(* Logix 5000 project; controller R400_500_XLS vendor 1 type 14 code 216 rev 31.11; software revision 31.01; part 20 of 32 *)
(* tags used below, declared in another part *)
   Alarm : SINT;   // Wait 3 seconds
   AlarmAcked : BOOL;   // Alarm has been acked
   AlarmFlag : DINT;   // Active alarm flag
   AlarmFlag1 : DINT;
   AlarmMuted : BOOL;
   AlarmTran0 : BOOL;   // Transition from step 3 to step 0
   Ashutdown : SINT;   // Not Used
   bAlrm : BOOL[64];
   Critical_Alarm : BOOL;
   CycExcBuffer : UDT_CYCLE;
   F2rinse : DINT;   // Not Used
   F3rinse : DINT;   // Not Used
   FC45_NextMaintDate : DINT[3];   // Next maintenance due date
   FINALRINSE_1 : DINT;   // Final rinse 1 id number
   HeatSmp : DINT;
   I_0_Missing : BOOL;
   L310ER_Led : DINT;
   LowPressAlmSp : REAL;   // Pump pressure too low setpoint
   M : DINT[5];   // Memory Bits
   ONS_FC45 : DINT;
   PWTnkTempAlmSp : REAL;   // Pure water tank temperature too high setpoint
   ResetMute : BOOL;
   Run : DINT;
   SumpTempAlmSp : REAL;   // Sump temperature too high setpoint
   Supervisor : DINT;
   Tmr : TIMER[107];
   Trt_Wsh : DINT;
   AlarmAck : INT;   // Alarm acknowledgement from the HMI
   AlarmTrigger : INT;   // Triggers the alarm screen if different of 0
   BatteryLowWarning : BOOL;
   bONSAuditTrailAlarm : BOOL;
   Current_Screen : DINT;
   DateTime : DINT[7];
   FC45_NbCycBeforeMaint : DINT;
   I_Ld_Dr_Cls_Sw : BOOL;   // Load door close
   I_MCR : BOOL;   // MCR input
   I_Mtr_Ovrld : BOOL;   // Motor overload
   I_Pw_Tnk_Sft_Lvl_Sw : BOOL;   // Pure water tank safety level switch
   I_Smp_Sft_Lvl_Sw : BOOL;   // Sump safety level switch
   I_Unld_Dr_Cls_Sw : BOOL;   // Unload door close
   I_UnldDr_ClseSlnce_Bttn : BOOL;   // Door Close/ Silence button Unload Side
   LastRecircSumpDrainTemp : REAL;
   Load : Doors;
   LoadDoorClosing : BOOL;
   LoadDoorOpening : BOOL;
   PmpPres : REAL;
   PureWaterTankTemp : REAL;   // Pure water tank temperature
   PWT_DeltaTempNeg : REAL;
   PWT_DeltaTempPos : REAL;
   Screen_Ctrl : DINT;   // PLC Screen Request
   SimGenEnabled : BOOL;   // SimGen enable bit 1= Simgen ON
   SPV_19 : BOOL;   // Screen 80 Enabled/Disabled Pump pressure monitoring
   SumpTemp : REAL;   // Sump temperature in °C
   tDelayBeforeFillingAuthAlarm : TIMER;
   tDelayBeforeTankFillingAuthAlarm : TIMER;
   Tpb : DINT[11];
   TreatmentPtr : DINT;
   udtAuditTrail : UDT_AuditTrail;
   Unit : Hrdwre;   // Unit Configuration
   UnLoad : Doors;
   UnloadDoorClosing : BOOL;
   UnloadDoorOpening : BOOL;
(* MainProgram, continued *)

ROUTINE WSH_10_WSH_37_GENERATE_ALARM_DISPLAY   (* ladder *)
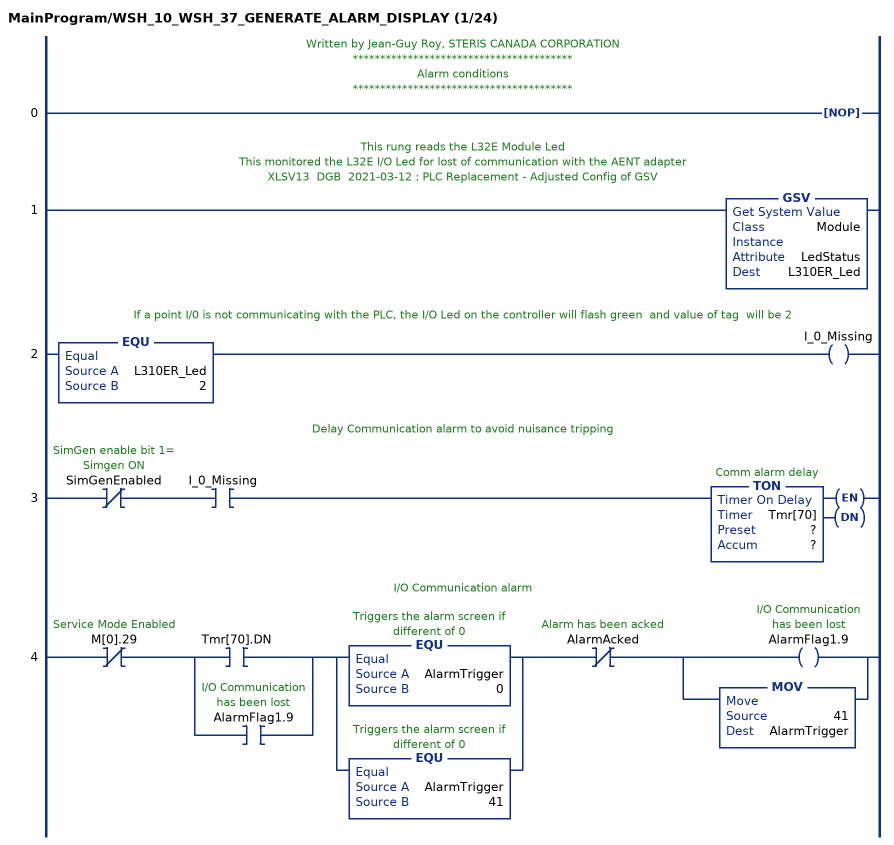
   // Written by Jean-Guy Roy, STERIS CANADA CORPORATION
   // ****************************************
   // Alarm conditions
   // ****************************************
   0: NOP();
   // This rung reads the L32E Module Led
   // This monitored the L32E I/O Led for lost of communication with the AENT adapter
   // XLSV13  DGB  2021-03-12 : PLC Replacement - Adjusted Config of GSV
   1: GSV(Module,,LedStatus,L310ER_Led);
   // If a point I/0 is not communicating with the PLC, the I/O Led on the controller will flash green  and value of tag  will be 2
   2: EQU(L310ER_Led,2)OTE(I_0_Missing);
   // Delay Communication alarm to avoid nuisance tripping
   3: XIO(SimGenEnabled)XIC(I_0_Missing)TON(Tmr[70],?,?);
   // I/O Communication alarm
   4: XIO(M[0].29)[XIC(Tmr[70].DN) ,XIC(AlarmFlag1.9) ][EQU(AlarmTrigger,0) ,EQU(AlarmTrigger,41) ]XIO(AlarmAcked)[OTE(AlarmFlag1.9) ,MOV(41,AlarmTrigger) ];
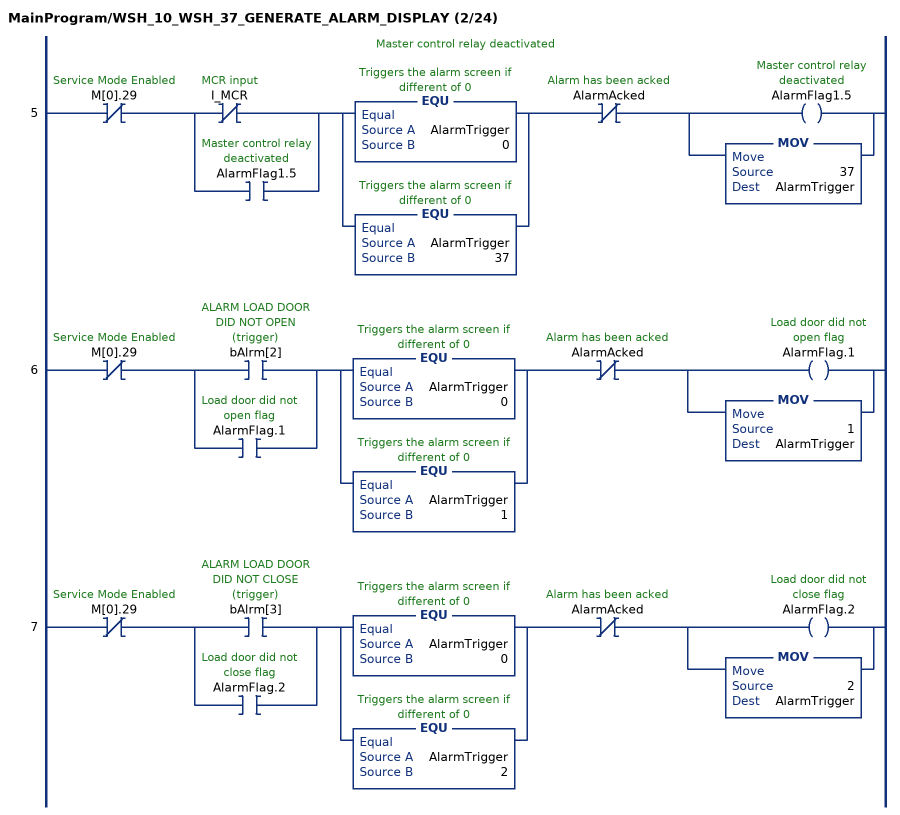
   // Master control relay deactivated
   5: XIO(M[0].29)[XIO(I_MCR) ,XIC(AlarmFlag1.5) ][EQU(AlarmTrigger,0) ,EQU(AlarmTrigger,37) ]XIO(AlarmAcked)[OTE(AlarmFlag1.5) ,MOV(37,AlarmTrigger) ];
   6: XIO(M[0].29)[XIC(bAlrm[2]) ,XIC(AlarmFlag.1) ][EQU(AlarmTrigger,0) ,EQU(AlarmTrigger,1) ]XIO(AlarmAcked)[OTE(AlarmFlag.1) ,MOV(1,AlarmTrigger) ];
   7: XIO(M[0].29)[XIC(bAlrm[3]) ,XIC(AlarmFlag.2) ][EQU(AlarmTrigger,0) ,EQU(AlarmTrigger,2) ]XIO(AlarmAcked)[OTE(AlarmFlag.2) ,MOV(2,AlarmTrigger) ];
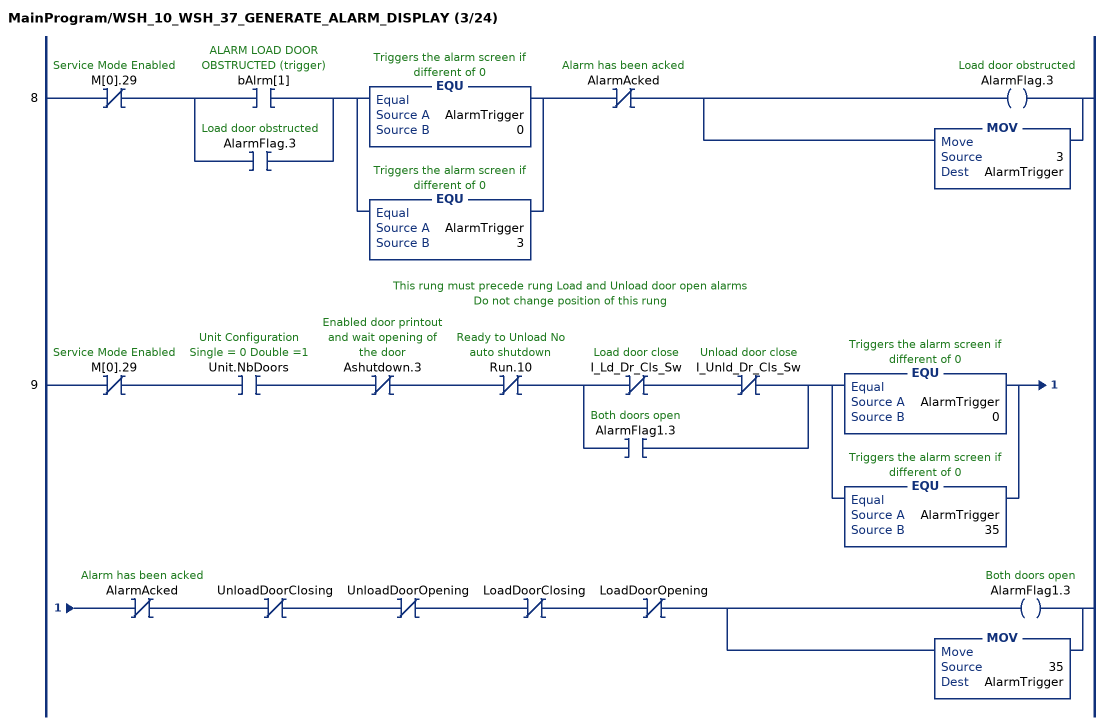
   8: XIO(M[0].29)[XIC(bAlrm[1]) ,XIC(AlarmFlag.3) ][EQU(AlarmTrigger,0) ,EQU(AlarmTrigger,3) ]XIO(AlarmAcked)[OTE(AlarmFlag.3) ,MOV(3,AlarmTrigger) ];
   // This rung must precede rung Load and Unload door open alarms
   // Do not change position of this rung
   9: XIO(M[0].29)XIC(Unit.NbDoors)XIO(Ashutdown.3)XIO(Run.10)[XIO(I_Ld_Dr_Cls_Sw) XIO(I_Unld_Dr_Cls_Sw) ,XIC(AlarmFlag1.3) ][EQU(AlarmTrigger,0) ,EQU(AlarmTrigger,35) ]XIO(AlarmAcked)XIO(UnloadDoorClosing)XIO(UnloadDoorOpening)XIO(LoadDoorClosing)XIO(LoadDoorOpening)[OTE(AlarmFlag1.3) ,MOV(35,AlarmTrigger) ];
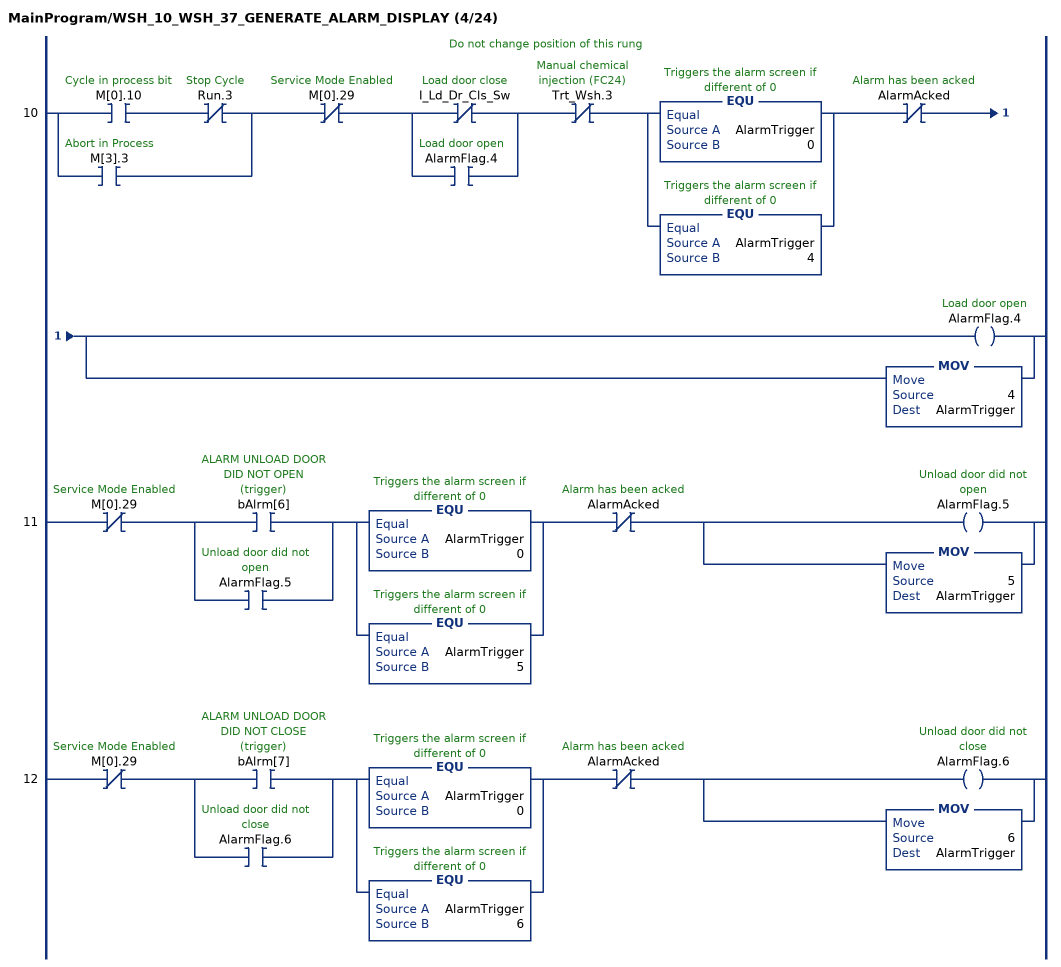
   // Do not change position of this rung
   10: [XIC(M[0].10) XIO(Run.3) ,XIC(M[3].3) ]XIO(M[0].29)[XIO(I_Ld_Dr_Cls_Sw) ,XIC(AlarmFlag.4) ]XIO(Trt_Wsh.3)[EQU(AlarmTrigger,0) ,EQU(AlarmTrigger,4) ]XIO(AlarmAcked)[OTE(AlarmFlag.4) ,MOV(4,AlarmTrigger) ];
   11: XIO(M[0].29)[XIC(bAlrm[6]) ,XIC(AlarmFlag.5) ][EQU(AlarmTrigger,0) ,EQU(AlarmTrigger,5) ]XIO(AlarmAcked)[OTE(AlarmFlag.5) ,MOV(5,AlarmTrigger) ];
   12: XIO(M[0].29)[XIC(bAlrm[7]) ,XIC(AlarmFlag.6) ][EQU(AlarmTrigger,0) ,EQU(AlarmTrigger,6) ]XIO(AlarmAcked)[OTE(AlarmFlag.6) ,MOV(6,AlarmTrigger) ];
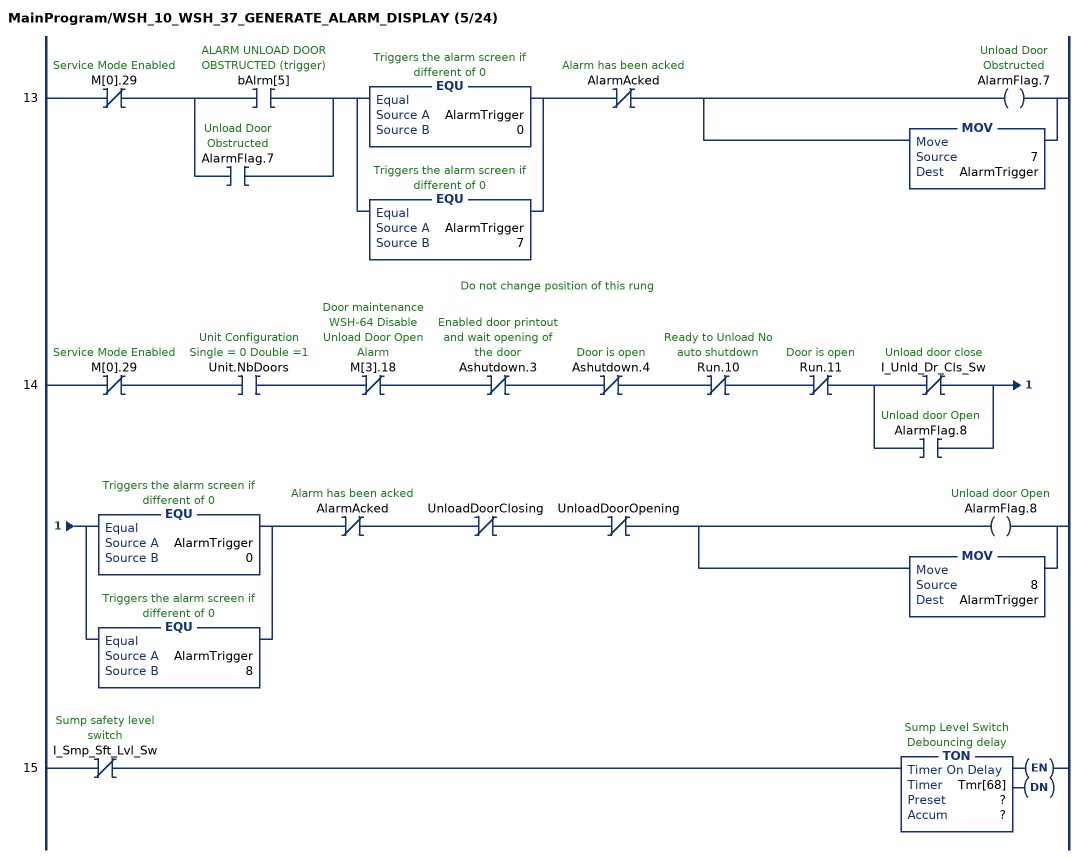
   13: XIO(M[0].29)[XIC(bAlrm[5]) ,XIC(AlarmFlag.7) ][EQU(AlarmTrigger,0) ,EQU(AlarmTrigger,7) ]XIO(AlarmAcked)[OTE(AlarmFlag.7) ,MOV(7,AlarmTrigger) ];
   // Do not change position of this rung
   14: XIO(M[0].29)XIC(Unit.NbDoors)XIO(M[3].18)XIO(Ashutdown.3)XIO(Ashutdown.4)XIO(Run.10)XIO(Run.11)[XIO(I_Unld_Dr_Cls_Sw) ,XIC(AlarmFlag.8) ][EQU(AlarmTrigger,0) ,EQU(AlarmTrigger,8) ]XIO(AlarmAcked)XIO(UnloadDoorClosing)XIO(UnloadDoorOpening)[OTE(AlarmFlag.8) ,MOV(8,AlarmTrigger) ];
   15: XIO(I_Smp_Sft_Lvl_Sw)TON(Tmr[68],?,?);
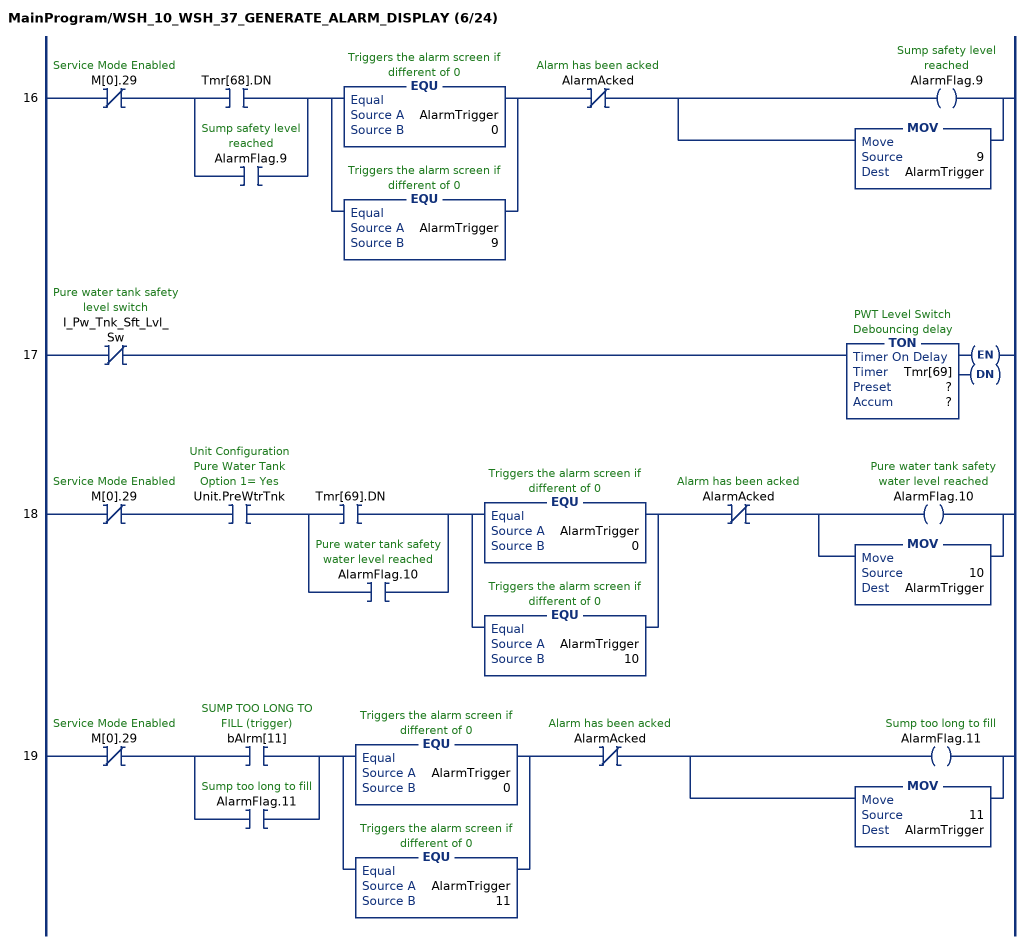
   16: XIO(M[0].29)[XIC(Tmr[68].DN) ,XIC(AlarmFlag.9) ][EQU(AlarmTrigger,0) ,EQU(AlarmTrigger,9) ]XIO(AlarmAcked)[OTE(AlarmFlag.9) ,MOV(9,AlarmTrigger) ];
   17: XIO(I_Pw_Tnk_Sft_Lvl_Sw)TON(Tmr[69],?,?);
   18: XIO(M[0].29)XIC(Unit.PreWtrTnk)[XIC(Tmr[69].DN) ,XIC(AlarmFlag.10) ][EQU(AlarmTrigger,0) ,EQU(AlarmTrigger,10) ]XIO(AlarmAcked)[OTE(AlarmFlag.10) ,MOV(10,AlarmTrigger) ];
   19: XIO(M[0].29)[XIC(bAlrm[11]) ,XIC(AlarmFlag.11) ][EQU(AlarmTrigger,0) ,EQU(AlarmTrigger,11) ]XIO(AlarmAcked)[OTE(AlarmFlag.11) ,MOV(11,AlarmTrigger) ];
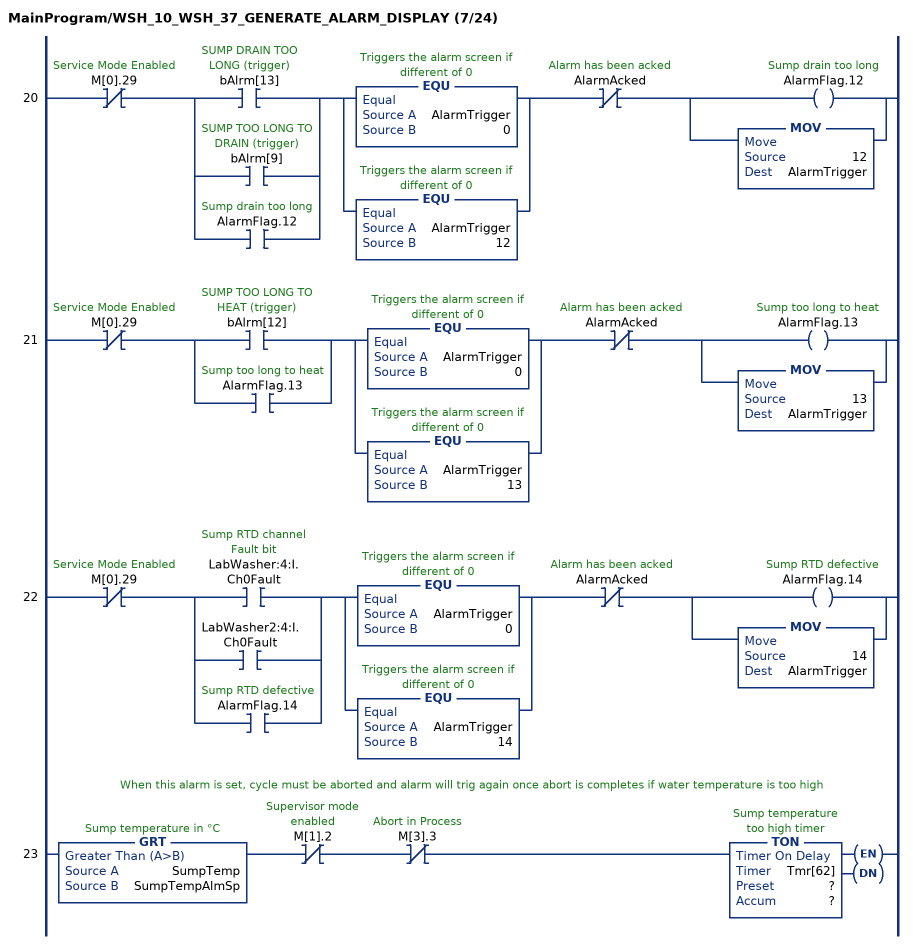
   20: XIO(M[0].29)[XIC(bAlrm[13]) ,XIC(bAlrm[9]) ,XIC(AlarmFlag.12) ][EQU(AlarmTrigger,0) ,EQU(AlarmTrigger,12) ]XIO(AlarmAcked)[OTE(AlarmFlag.12) ,MOV(12,AlarmTrigger) ];
   21: XIO(M[0].29)[XIC(bAlrm[12]) ,XIC(AlarmFlag.13) ][EQU(AlarmTrigger,0) ,EQU(AlarmTrigger,13) ]XIO(AlarmAcked)[OTE(AlarmFlag.13) ,MOV(13,AlarmTrigger) ];
   22: XIO(M[0].29)[XIC(LabWasher:4:I.Ch0Fault) ,XIC(LabWasher2:4:I.Ch0Fault) ,XIC(AlarmFlag.14) ][EQU(AlarmTrigger,0) ,EQU(AlarmTrigger,14) ]XIO(AlarmAcked)[OTE(AlarmFlag.14) ,MOV(14,AlarmTrigger) ];
   // When this alarm is set, cycle must be aborted and alarm will trig again once abort is completes if water temperature is too high
   23: GRT(SumpTemp,SumpTempAlmSp)XIO(M[1].2)XIO(M[3].3)TON(Tmr[62],?,?);
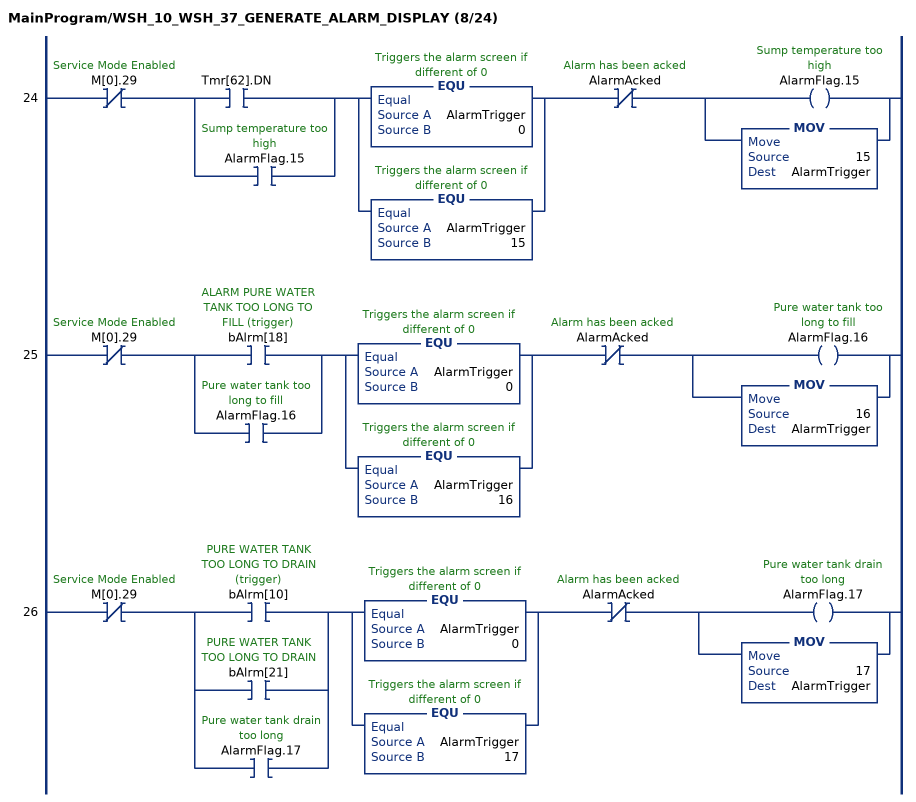
   24: XIO(M[0].29)[XIC(Tmr[62].DN) ,XIC(AlarmFlag.15) ][EQU(AlarmTrigger,0) ,EQU(AlarmTrigger,15) ]XIO(AlarmAcked)[OTE(AlarmFlag.15) ,MOV(15,AlarmTrigger) ];
   25: XIO(M[0].29)[XIC(bAlrm[18]) ,XIC(AlarmFlag.16) ][EQU(AlarmTrigger,0) ,EQU(AlarmTrigger,16) ]XIO(AlarmAcked)[OTE(AlarmFlag.16) ,MOV(16,AlarmTrigger) ];
   26: XIO(M[0].29)[XIC(bAlrm[10]) ,XIC(bAlrm[21]) ,XIC(AlarmFlag.17) ][EQU(AlarmTrigger,0) ,EQU(AlarmTrigger,17) ]XIO(AlarmAcked)[OTE(AlarmFlag.17) ,MOV(17,AlarmTrigger) ];
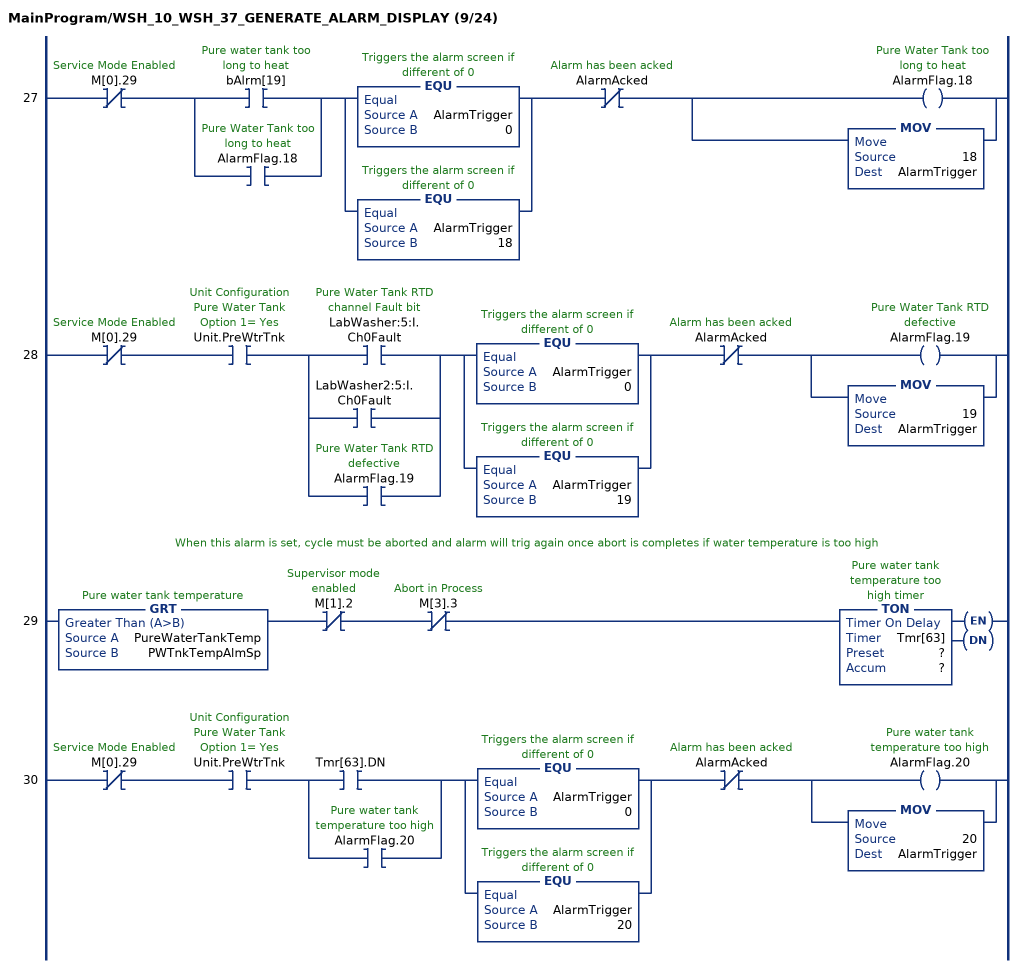
   27: XIO(M[0].29)[XIC(bAlrm[19]) ,XIC(AlarmFlag.18) ][EQU(AlarmTrigger,0) ,EQU(AlarmTrigger,18) ]XIO(AlarmAcked)[OTE(AlarmFlag.18) ,MOV(18,AlarmTrigger) ];
   28: XIO(M[0].29)XIC(Unit.PreWtrTnk)[XIC(LabWasher:5:I.Ch0Fault) ,XIC(LabWasher2:5:I.Ch0Fault) ,XIC(AlarmFlag.19) ][EQU(AlarmTrigger,0) ,EQU(AlarmTrigger,19) ]XIO(AlarmAcked)[OTE(AlarmFlag.19) ,MOV(19,AlarmTrigger) ];
   // When this alarm is set, cycle must be aborted and alarm will trig again once abort is completes if water temperature is too high
   29: GRT(PureWaterTankTemp,PWTnkTempAlmSp)XIO(M[1].2)XIO(M[3].3)TON(Tmr[63],?,?);
   30: XIO(M[0].29)XIC(Unit.PreWtrTnk)[XIC(Tmr[63].DN) ,XIC(AlarmFlag.20) ][EQU(AlarmTrigger,0) ,EQU(AlarmTrigger,20) ]XIO(AlarmAcked)[OTE(AlarmFlag.20) ,MOV(20,AlarmTrigger) ];
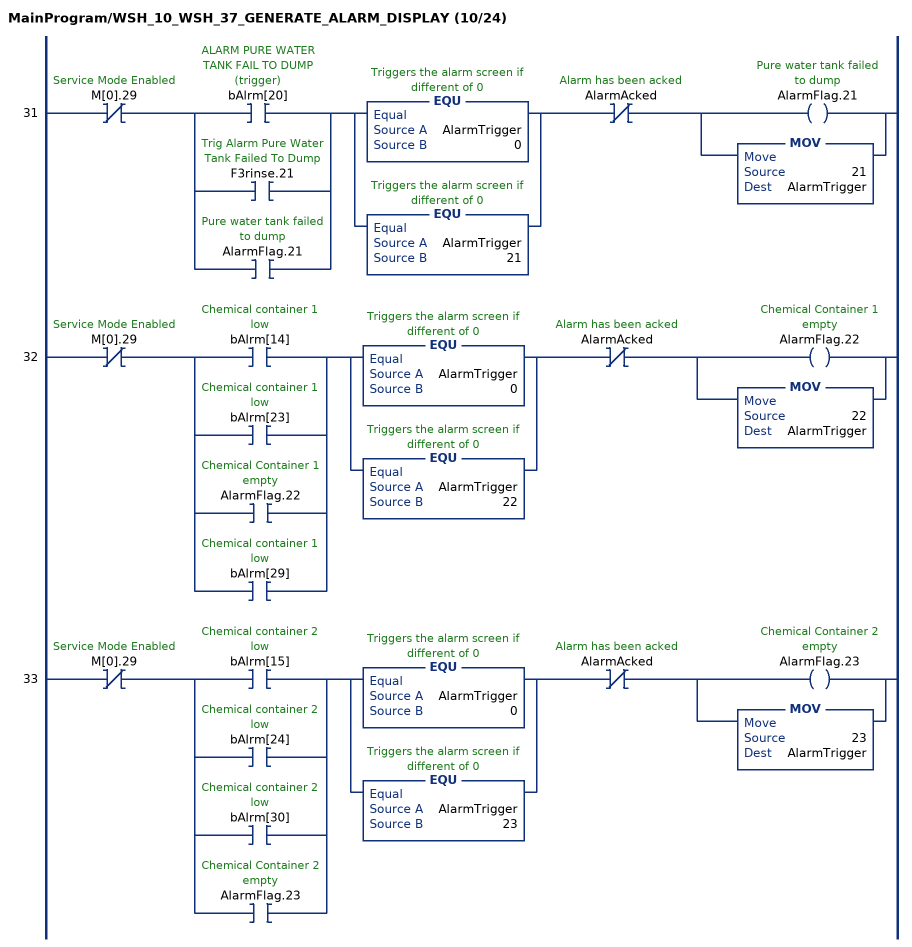
   31: XIO(M[0].29)[XIC(bAlrm[20]) ,XIC(F3rinse.21) ,XIC(AlarmFlag.21) ][EQU(AlarmTrigger,0) ,EQU(AlarmTrigger,21) ]XIO(AlarmAcked)[OTE(AlarmFlag.21) ,MOV(21,AlarmTrigger) ];
   32: XIO(M[0].29)[XIC(bAlrm[14]) ,XIC(bAlrm[23]) ,XIC(AlarmFlag.22) ,XIC(bAlrm[29]) ][EQU(AlarmTrigger,0) ,EQU(AlarmTrigger,22) ]XIO(AlarmAcked)[OTE(AlarmFlag.22) ,MOV(22,AlarmTrigger) ];
   33: XIO(M[0].29)[XIC(bAlrm[15]) ,XIC(bAlrm[24]) ,XIC(bAlrm[30]) ,XIC(AlarmFlag.23) ][EQU(AlarmTrigger,0) ,EQU(AlarmTrigger,23) ]XIO(AlarmAcked)[OTE(AlarmFlag.23) ,MOV(23,AlarmTrigger) ];
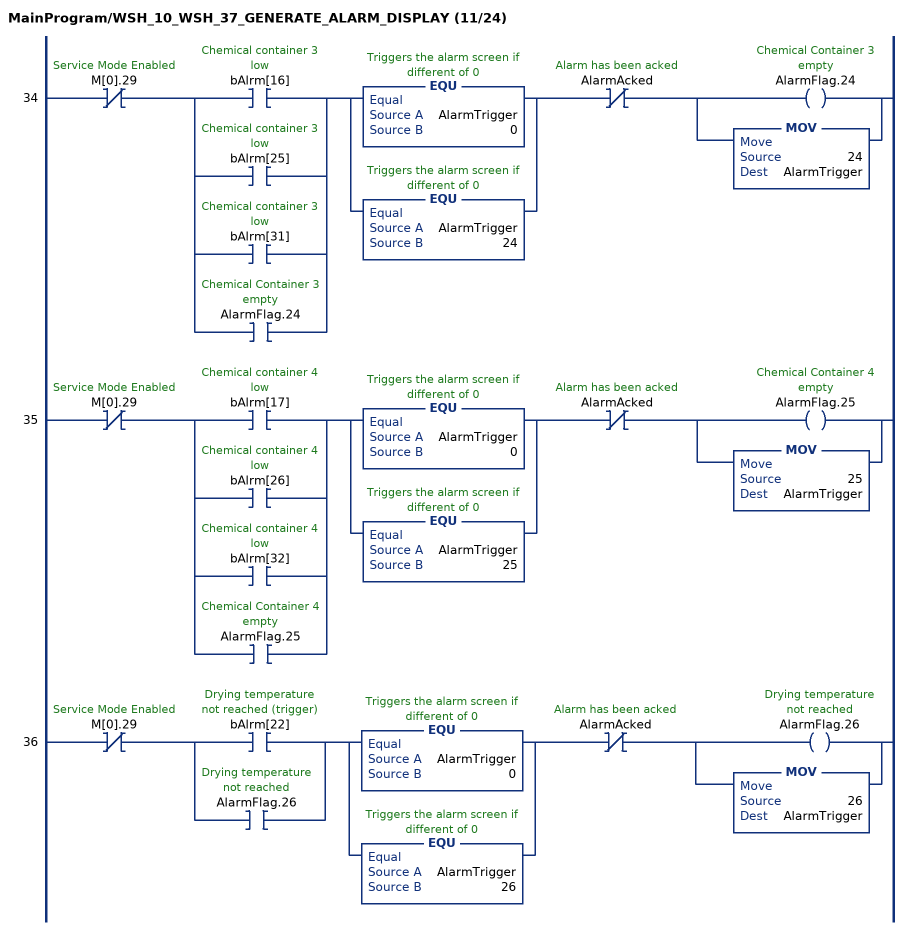
   34: XIO(M[0].29)[XIC(bAlrm[16]) ,XIC(bAlrm[25]) ,XIC(bAlrm[31]) ,XIC(AlarmFlag.24) ][EQU(AlarmTrigger,0) ,EQU(AlarmTrigger,24) ]XIO(AlarmAcked)[OTE(AlarmFlag.24) ,MOV(24,AlarmTrigger) ];
   35: XIO(M[0].29)[XIC(bAlrm[17]) ,XIC(bAlrm[26]) ,XIC(bAlrm[32]) ,XIC(AlarmFlag.25) ][EQU(AlarmTrigger,0) ,EQU(AlarmTrigger,25) ]XIO(AlarmAcked)[OTE(AlarmFlag.25) ,MOV(25,AlarmTrigger) ];
   36: XIO(M[0].29)[XIC(bAlrm[22]) ,XIC(AlarmFlag.26) ][EQU(AlarmTrigger,0) ,EQU(AlarmTrigger,26) ]XIO(AlarmAcked)[OTE(AlarmFlag.26) ,MOV(26,AlarmTrigger) ];
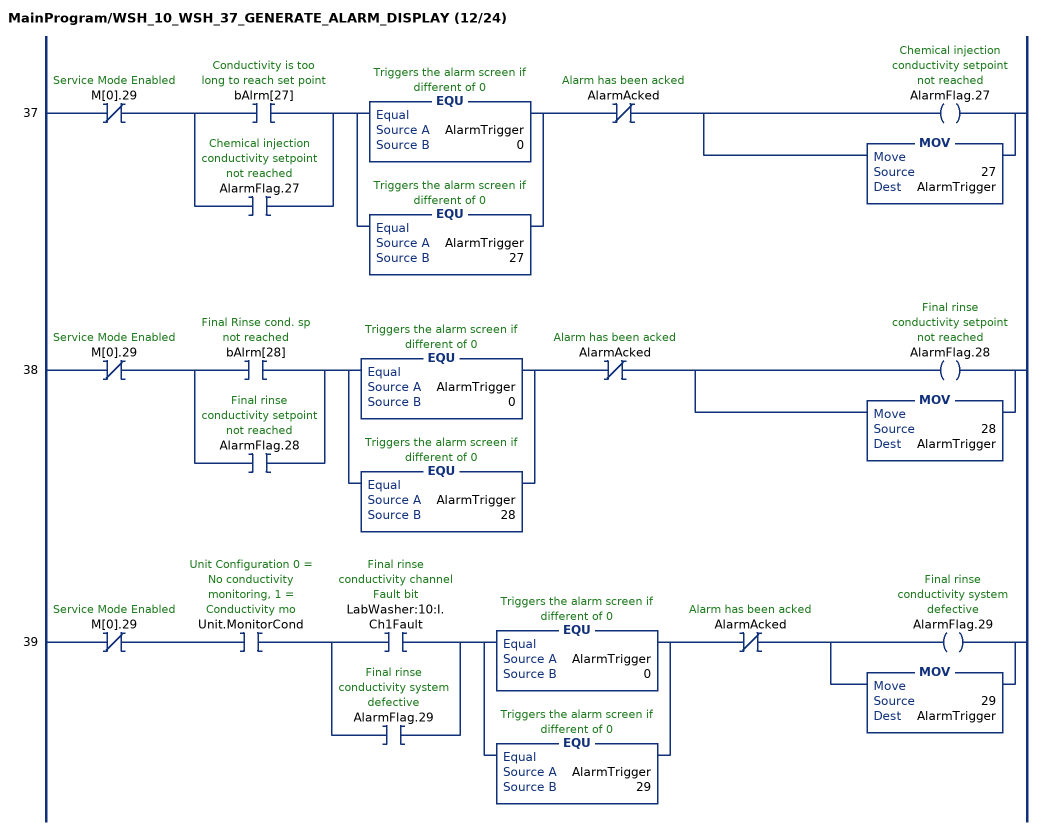
   37: XIO(M[0].29)[XIC(bAlrm[27]) ,XIC(AlarmFlag.27) ][EQU(AlarmTrigger,0) ,EQU(AlarmTrigger,27) ]XIO(AlarmAcked)[OTE(AlarmFlag.27) ,MOV(27,AlarmTrigger) ];
   38: XIO(M[0].29)[XIC(bAlrm[28]) ,XIC(AlarmFlag.28) ][EQU(AlarmTrigger,0) ,EQU(AlarmTrigger,28) ]XIO(AlarmAcked)[OTE(AlarmFlag.28) ,MOV(28,AlarmTrigger) ];
   39: XIO(M[0].29)XIC(Unit.MonitorCond)[XIC(LabWasher:10:I.Ch1Fault) ,XIC(AlarmFlag.29) ][EQU(AlarmTrigger,0) ,EQU(AlarmTrigger,29) ]XIO(AlarmAcked)[OTE(AlarmFlag.29) ,MOV(29,AlarmTrigger) ];
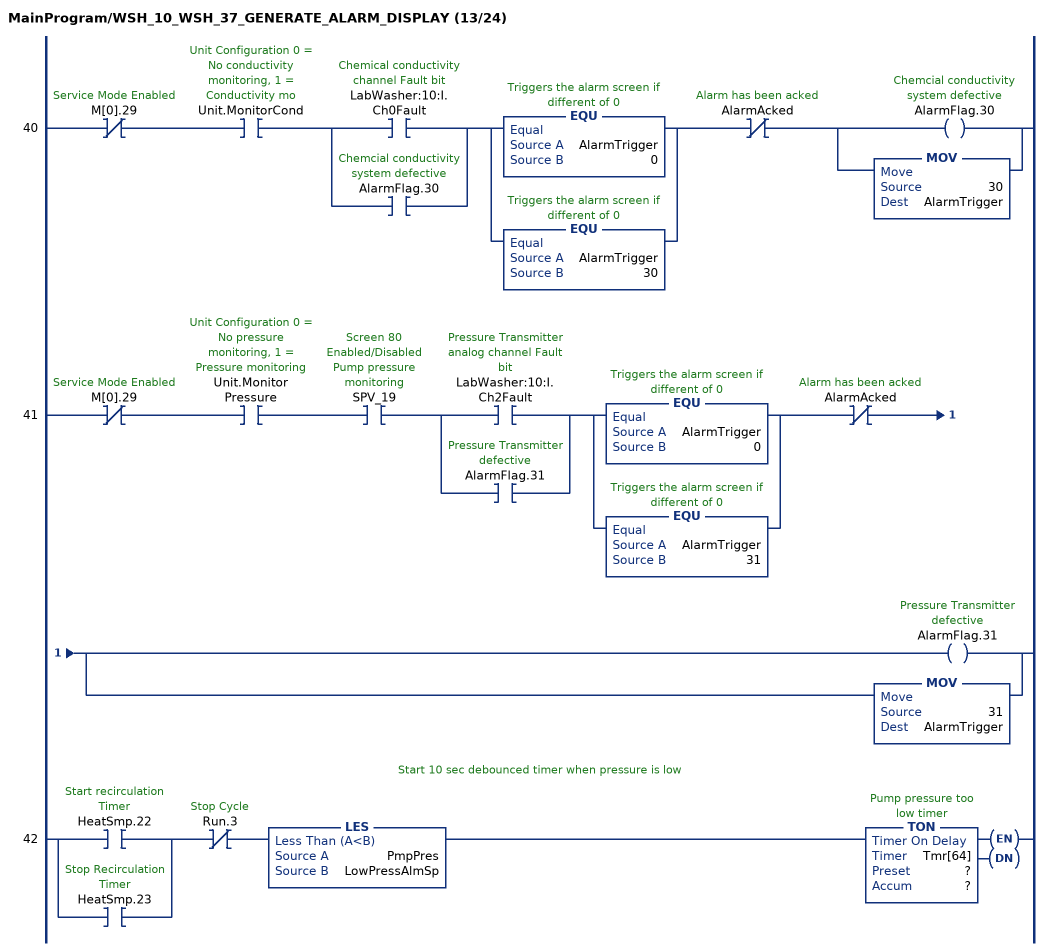
   40: XIO(M[0].29)XIC(Unit.MonitorCond)[XIC(LabWasher:10:I.Ch0Fault) ,XIC(AlarmFlag.30) ][EQU(AlarmTrigger,0) ,EQU(AlarmTrigger,30) ]XIO(AlarmAcked)[OTE(AlarmFlag.30) ,MOV(30,AlarmTrigger) ];
   41: XIO(M[0].29)XIC(Unit.MonitorPressure)XIC(SPV_19)[XIC(LabWasher:10:I.Ch2Fault) ,XIC(AlarmFlag.31) ][EQU(AlarmTrigger,0) ,EQU(AlarmTrigger,31) ]XIO(AlarmAcked)[OTE(AlarmFlag.31) ,MOV(31,AlarmTrigger) ];
   // Start 10 sec debounced timer when pressure is low
   42: [XIC(HeatSmp.22) ,XIC(HeatSmp.23) ]XIO(Run.3)LES(PmpPres,LowPressAlmSp)TON(Tmr[64],?,?);
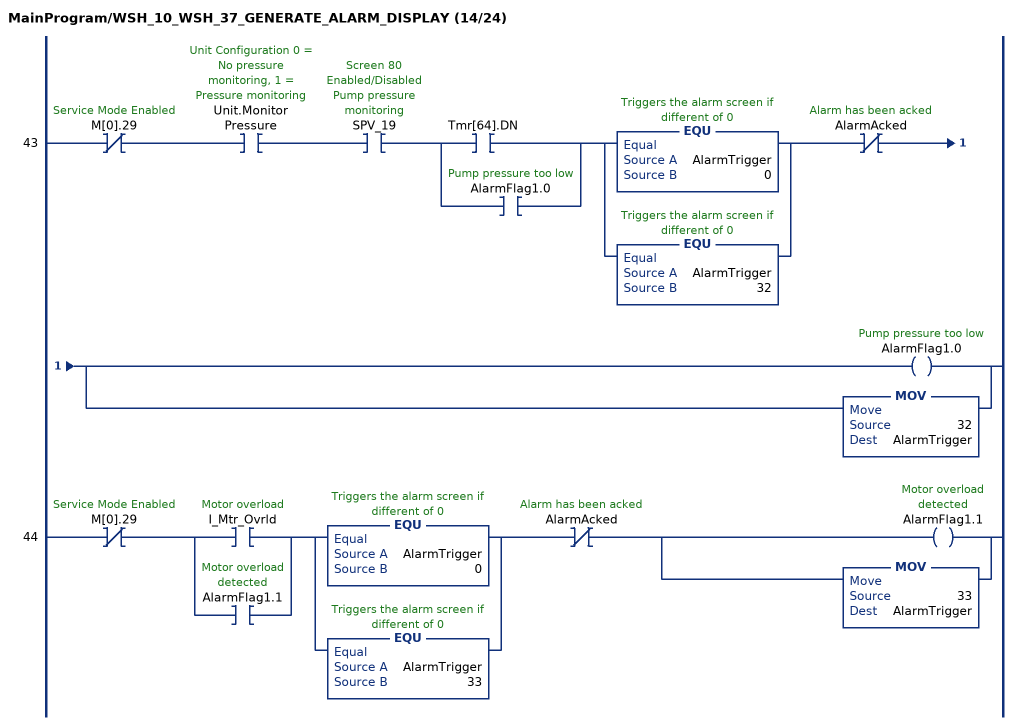
   43: XIO(M[0].29)XIC(Unit.MonitorPressure)XIC(SPV_19)[XIC(Tmr[64].DN) ,XIC(AlarmFlag1.0) ][EQU(AlarmTrigger,0) ,EQU(AlarmTrigger,32) ]XIO(AlarmAcked)[OTE(AlarmFlag1.0) ,MOV(32,AlarmTrigger) ];
   44: XIO(M[0].29)[XIC(I_Mtr_Ovrld) ,XIC(AlarmFlag1.1) ][EQU(AlarmTrigger,0) ,EQU(AlarmTrigger,33) ]XIO(AlarmAcked)[OTE(AlarmFlag1.1) ,MOV(33,AlarmTrigger) ];
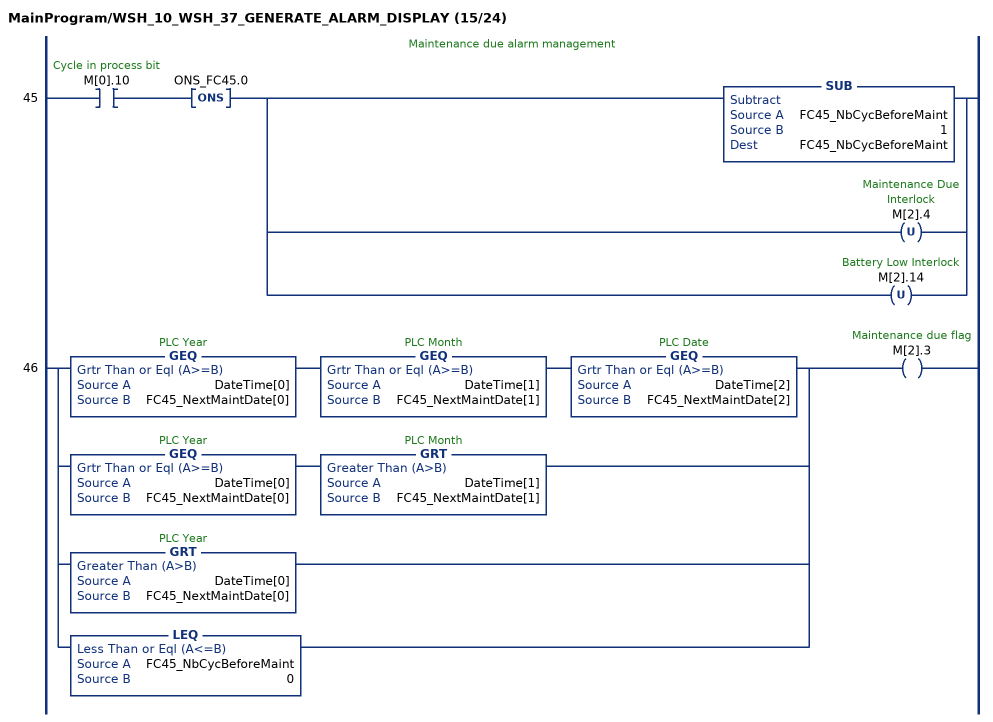
   // Maintenance due alarm management
   45: XIC(M[0].10)ONS(ONS_FC45.0)[SUB(FC45_NbCycBeforeMaint,1,FC45_NbCycBeforeMaint) ,OTU(M[2].4) ,OTU(M[2].14) ];
   46: [GEQ(DateTime[0],FC45_NextMaintDate[0]) GEQ(DateTime[1],FC45_NextMaintDate[1]) GEQ(DateTime[2],FC45_NextMaintDate[2]) ,GEQ(DateTime[0],FC45_NextMaintDate[0]) GRT(DateTime[1],FC45_NextMaintDate[1]) ,GRT(DateTime[0],FC45_NextMaintDate[0]) ,LEQ(FC45_NbCycBeforeMaint,0) ]OTE(M[2].3);
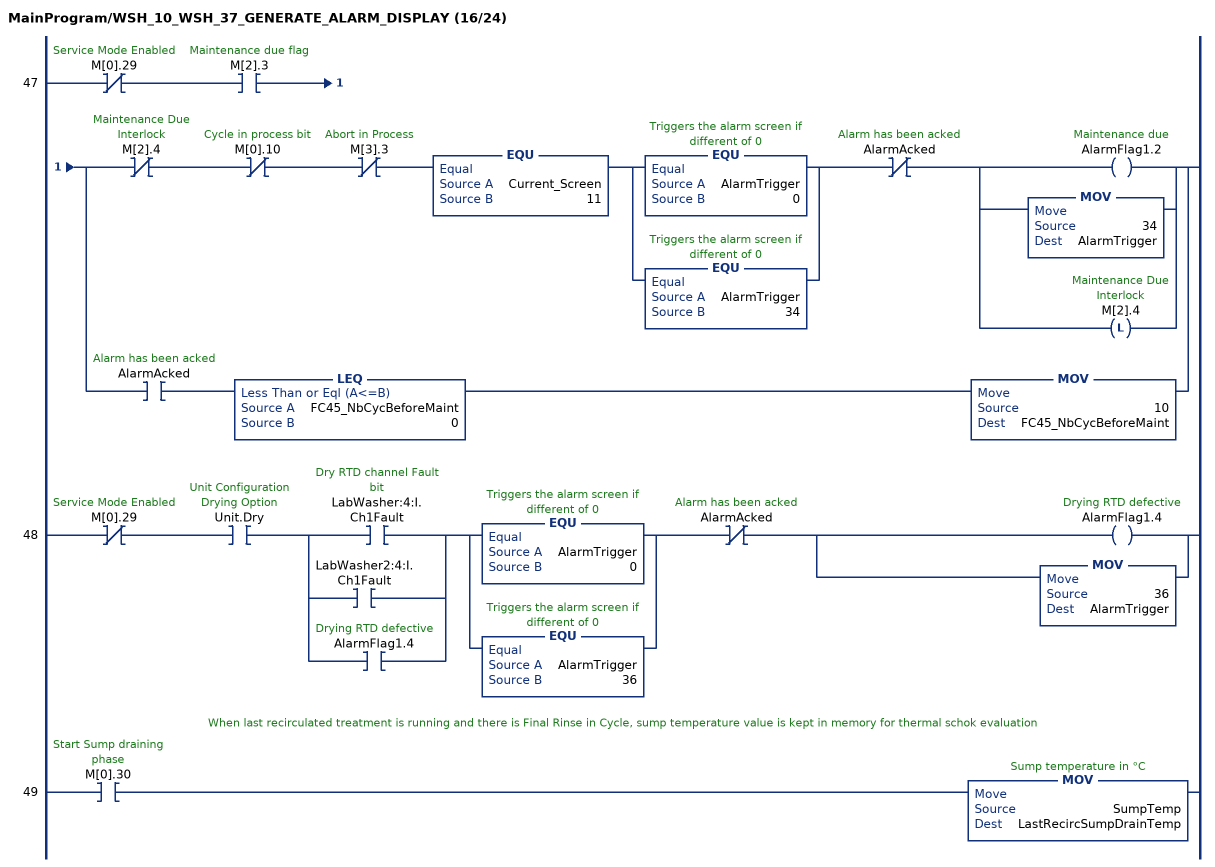
   47: XIO(M[0].29)XIC(M[2].3)[XIO(M[2].4) XIO(M[0].10) XIO(M[3].3) EQU(Current_Screen,11) [EQU(AlarmTrigger,0) ,EQU(AlarmTrigger,34) ] XIO(AlarmAcked) [OTE(AlarmFlag1.2) ,MOV(34,AlarmTrigger) ,OTL(M[2].4) ] ,XIC(AlarmAcked) LEQ(FC45_NbCycBeforeMaint,0) MOV(10,FC45_NbCycBeforeMaint) ];
   48: XIO(M[0].29)XIC(Unit.Dry)[XIC(LabWasher:4:I.Ch1Fault) ,XIC(LabWasher2:4:I.Ch1Fault) ,XIC(AlarmFlag1.4) ][EQU(AlarmTrigger,0) ,EQU(AlarmTrigger,36) ]XIO(AlarmAcked)[OTE(AlarmFlag1.4) ,MOV(36,AlarmTrigger) ];
   // When last recirculated treatment is running and there is Final Rinse in Cycle, sump temperature value is kept in memory for thermal schok evaluation
   49: XIC(M[0].30)MOV(SumpTemp,LastRecircSumpDrainTemp);
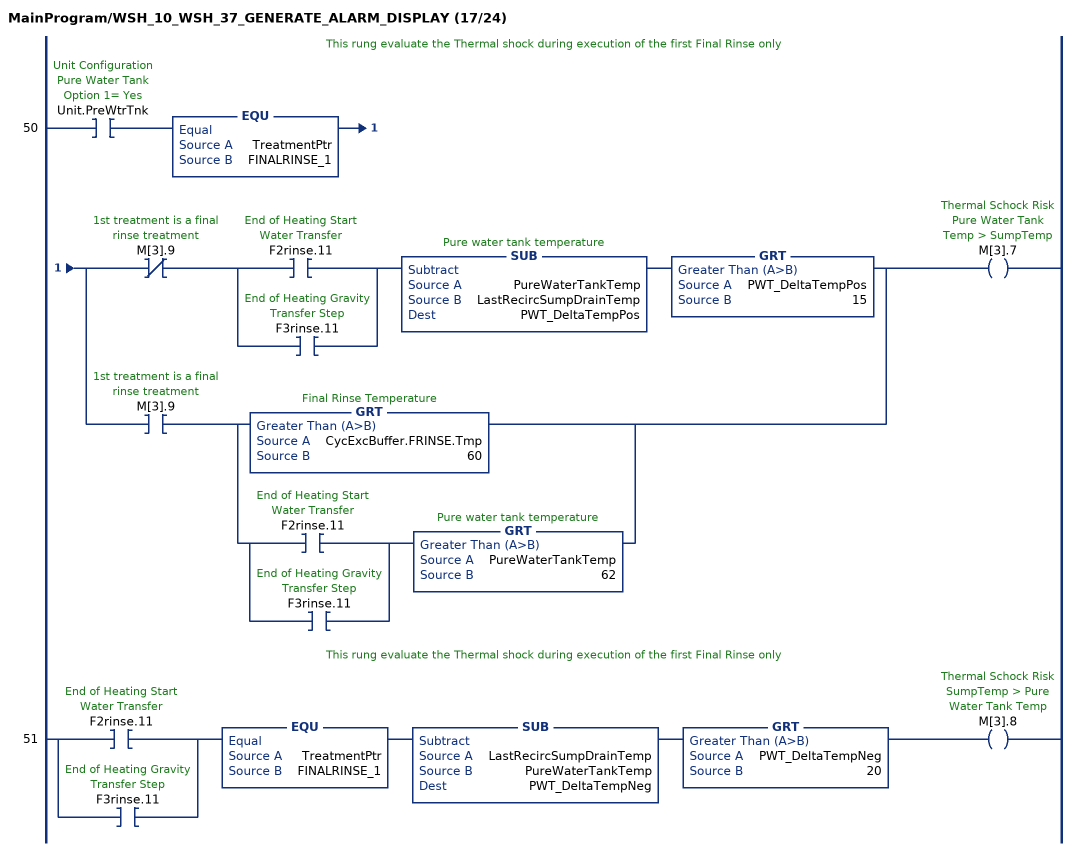
   // This rung evaluate the Thermal shock during execution of the first Final Rinse only
   50: XIC(Unit.PreWtrTnk)EQU(TreatmentPtr,FINALRINSE_1)[XIO(M[3].9) [XIC(F2rinse.11) ,XIC(F3rinse.11) ] SUB(PureWaterTankTemp,LastRecircSumpDrainTemp,PWT_DeltaTempPos) GRT(PWT_DeltaTempPos,15) ,XIC(M[3].9) [GRT(CycExcBuffer.FRINSE.Tmp,60) ,[XIC(F2rinse.11) ,XIC(F3rinse.11) ] GRT(PureWaterTankTemp,62) ] ]OTE(M[3].7);
   // This rung evaluate the Thermal shock during execution of the first Final Rinse only
   51: [XIC(F2rinse.11) ,XIC(F3rinse.11) ]EQU(TreatmentPtr,FINALRINSE_1)SUB(LastRecircSumpDrainTemp,PureWaterTankTemp,PWT_DeltaTempNeg)GRT(PWT_DeltaTempNeg,20)OTE(M[3].8);
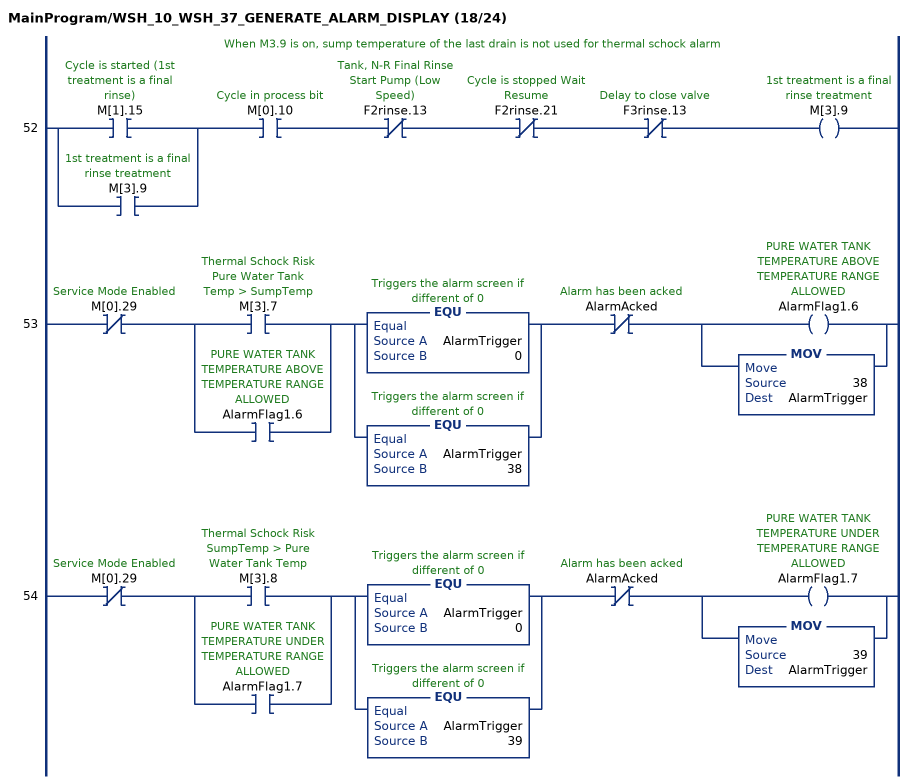
   // When M3.9 is on, sump temperature of the last drain is not used for thermal schock alarm
   52: [XIC(M[1].15) ,XIC(M[3].9) ]XIC(M[0].10)XIO(F2rinse.13)XIO(F2rinse.21)XIO(F3rinse.13)OTE(M[3].9);
   53: XIO(M[0].29)[XIC(M[3].7) ,XIC(AlarmFlag1.6) ][EQU(AlarmTrigger,0) ,EQU(AlarmTrigger,38) ]XIO(AlarmAcked)[OTE(AlarmFlag1.6) ,MOV(38,AlarmTrigger) ];
   54: XIO(M[0].29)[XIC(M[3].8) ,XIC(AlarmFlag1.7) ][EQU(AlarmTrigger,0) ,EQU(AlarmTrigger,39) ]XIO(AlarmAcked)[OTE(AlarmFlag1.7) ,MOV(39,AlarmTrigger) ];
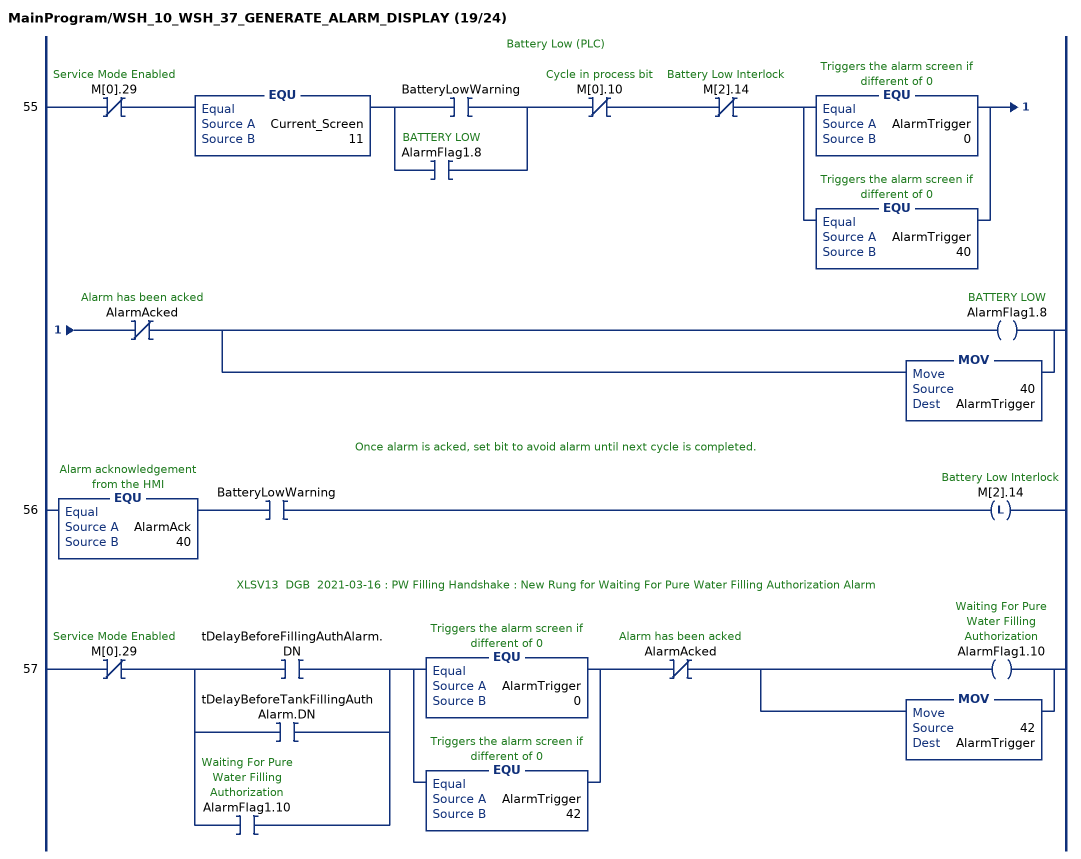
   // Battery Low (PLC)
   55: XIO(M[0].29)EQU(Current_Screen,11)[XIC(BatteryLowWarning) ,XIC(AlarmFlag1.8) ]XIO(M[0].10)XIO(M[2].14)[EQU(AlarmTrigger,0) ,EQU(AlarmTrigger,40) ]XIO(AlarmAcked)[OTE(AlarmFlag1.8) ,MOV(40,AlarmTrigger) ];
   // Once alarm is acked, set bit to avoid alarm until next cycle is completed.
   56: EQU(AlarmAck,40)XIC(BatteryLowWarning)OTL(M[2].14);
   // XLSV13  DGB  2021-03-16 : PW Filling Handshake : New Rung for Waiting For Pure Water Filling Authorization Alarm
   57: XIO(M[0].29)[XIC(tDelayBeforeFillingAuthAlarm.DN) ,XIC(tDelayBeforeTankFillingAuthAlarm.DN) ,XIC(AlarmFlag1.10) ][EQU(AlarmTrigger,0) ,EQU(AlarmTrigger,42) ]XIO(AlarmAcked)[OTE(AlarmFlag1.10) ,MOV(42,AlarmTrigger) ];
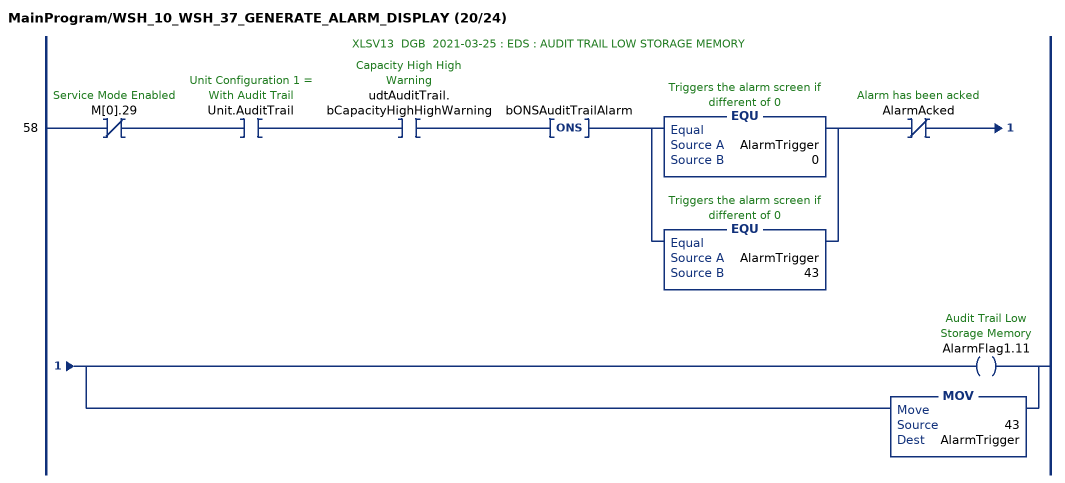
   // XLSV13  DGB  2021-03-25 : EDS : AUDIT TRAIL LOW STORAGE MEMORY
   58: XIO(M[0].29)XIC(Unit.AuditTrail)XIC(udtAuditTrail.bCapacityHighHighWarning)ONS(bONSAuditTrailAlarm)[EQU(AlarmTrigger,0) ,EQU(AlarmTrigger,43) ]XIO(AlarmAcked)[OTE(AlarmFlag1.11) ,MOV(43,AlarmTrigger) ];
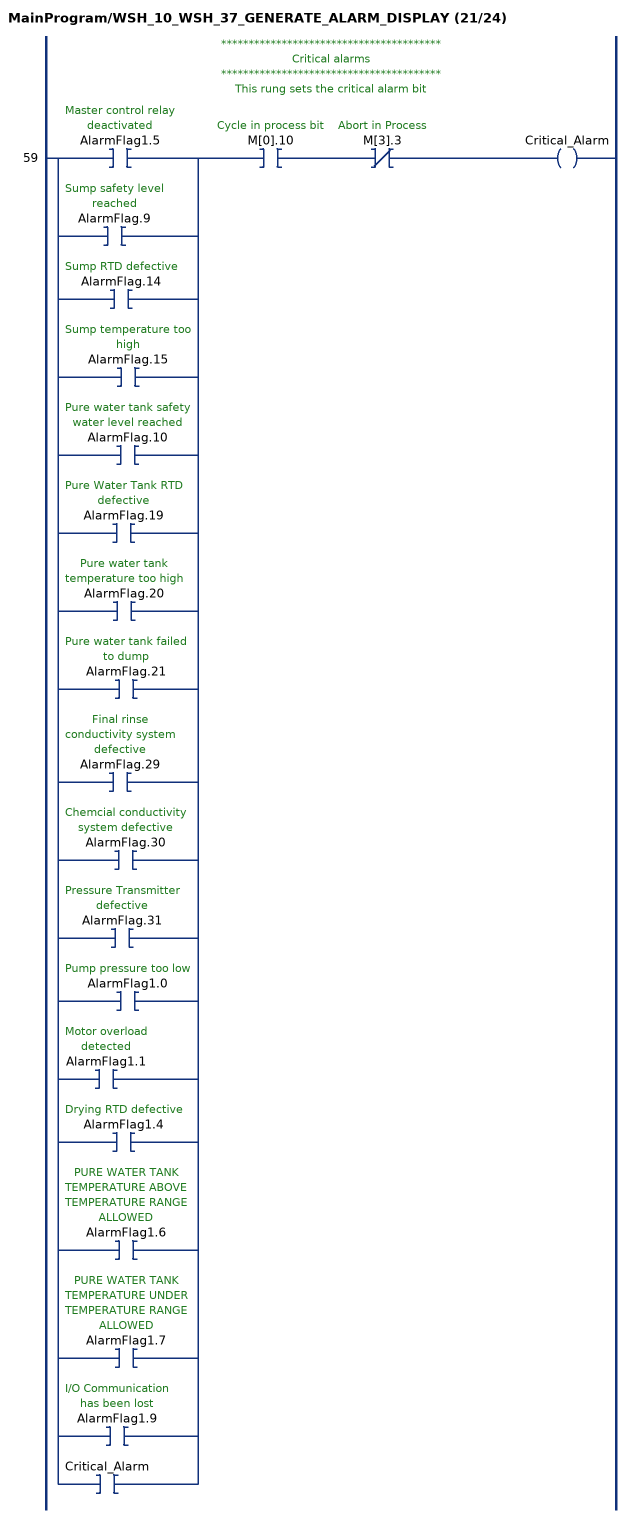
   // ****************************************
   // Critical alarms
   // ****************************************
   // This rung sets the critical alarm bit
   59: [XIC(AlarmFlag1.5) ,XIC(AlarmFlag.9) ,XIC(AlarmFlag.14) ,XIC(AlarmFlag.15) ,XIC(AlarmFlag.10) ,XIC(AlarmFlag.19) ,XIC(AlarmFlag.20) ,XIC(AlarmFlag.21) ,XIC(AlarmFlag.29) ,XIC(AlarmFlag.30) ,XIC(AlarmFlag.31) ,XIC(AlarmFlag1.0) ,XIC(AlarmFlag1.1) ,XIC(AlarmFlag1.4) ,XIC(AlarmFlag1.6) ,XIC(AlarmFlag1.7) ,XIC(AlarmFlag1.9) ,XIC(Critical_Alarm) ]XIC(M[0].10)XIO(M[3].3)OTE(Critical_Alarm);
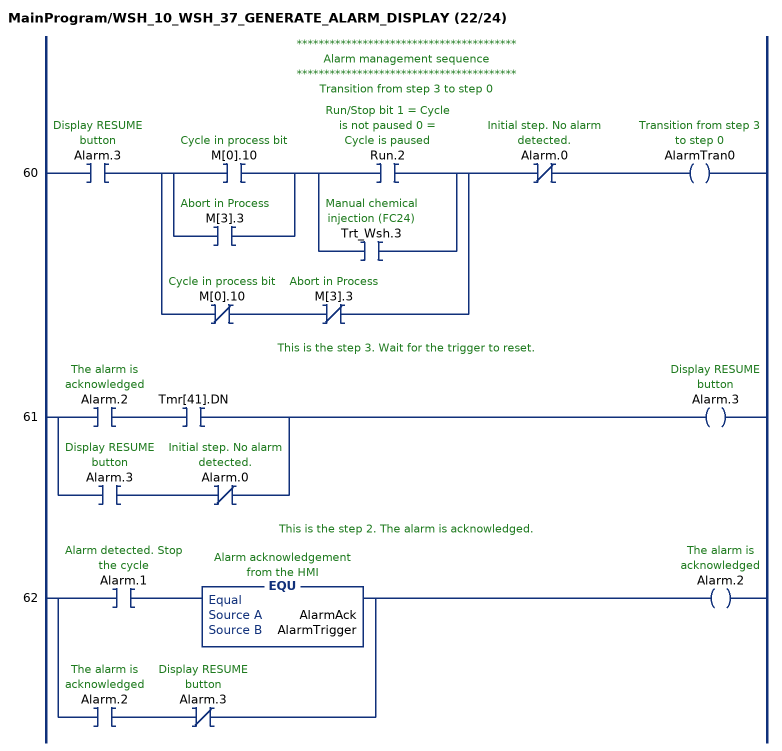
   // ****************************************
   // Alarm management sequence
   // ****************************************
   // Transition from step 3 to step 0
   60: XIC(Alarm.3)[[XIC(M[0].10) ,XIC(M[3].3) ] [XIC(Run.2) ,XIC(Trt_Wsh.3) ] ,XIO(M[0].10) XIO(M[3].3) ]XIO(Alarm.0)OTE(AlarmTran0);
   // This is the step 3. Wait for the trigger to reset.
   61: [XIC(Alarm.2) XIC(Tmr[41].DN) ,XIC(Alarm.3) XIO(Alarm.0) ]OTE(Alarm.3);
   // This is the step 2. The alarm is acknowledged.
   62: [XIC(Alarm.1) EQU(AlarmAck,AlarmTrigger) ,XIC(Alarm.2) XIO(Alarm.3) ]OTE(Alarm.2);
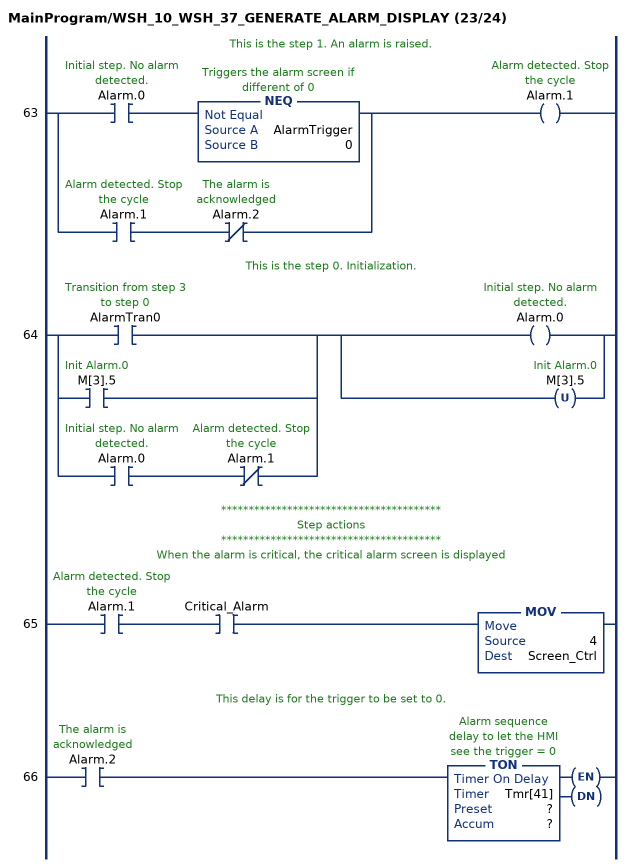
   // This is the step 1. An alarm is raised.
   63: [XIC(Alarm.0) NEQ(AlarmTrigger,0) ,XIC(Alarm.1) XIO(Alarm.2) ]OTE(Alarm.1);
   // This is the step 0. Initialization.
   64: [XIC(AlarmTran0) ,XIC(M[3].5) ,XIC(Alarm.0) XIO(Alarm.1) ][OTE(Alarm.0) ,OTU(M[3].5) ];
   // ****************************************
   // Step actions
   // ****************************************
   // When the alarm is critical, the critical alarm screen is displayed
   65: XIC(Alarm.1)XIC(Critical_Alarm)MOV(4,Screen_Ctrl);
   // This delay is for the trigger to be set to 0.
   66: XIC(Alarm.2)TON(Tmr[41],?,?);
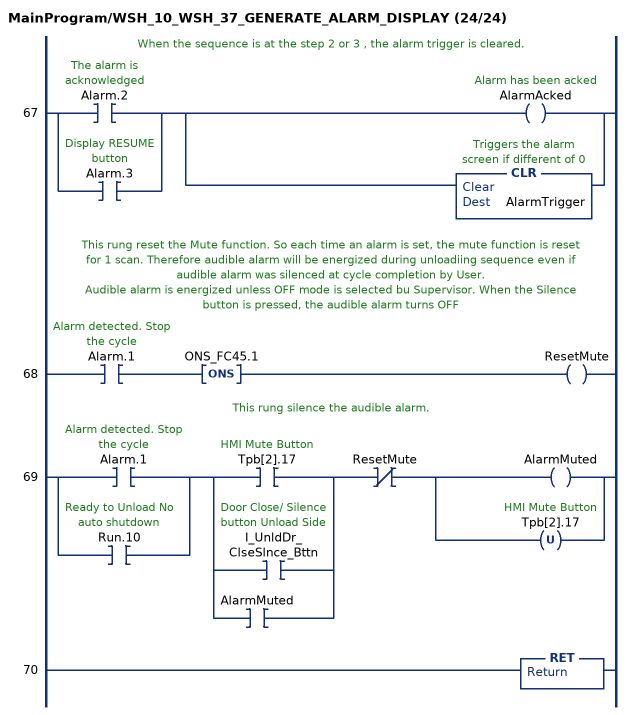
   // When the sequence is at the step 2 or 3 , the alarm trigger is cleared.
   67: [XIC(Alarm.2) ,XIC(Alarm.3) ][OTE(AlarmAcked) ,CLR(AlarmTrigger) ];
   // This rung reset the Mute function. So each time an alarm is set, the mute function is reset for 1 scan. Therefore audible alarm will be energized during unloadiing sequence even if audible alarm was silenced at cycle completion by User.
   // Audible alarm is energized unless OFF mode is selected bu Supervisor. When the Silence button is pressed, the audible alarm turns OFF
   68: XIC(Alarm.1)ONS(ONS_FC45.1)OTE(ResetMute);
   // This rung silence the audible alarm.
   69: [XIC(Alarm.1) ,XIC(Run.10) ][XIC(Tpb[2].17) ,XIC(I_UnldDr_ClseSlnce_Bttn) ,XIC(AlarmMuted) ]XIO(ResetMute)[OTE(AlarmMuted) ,OTU(Tpb[2].17) ];
   70: RET();
END_ROUTINE
